// TIA Portal V21 export
FUNCTION_BLOCK "FB_StarterStl"   // FB103, STL
TITLE = Пускатель насоса (STL)
{ S7_Optimized_Access := 'FALSE' }
AUTHOR : WTP2
FAMILY : Drives
VERSION : 0.1
// Пускатель насоса с контролем обратной связи (один блок на LAD, FBD, STL, SCL).
// 1. Пуск/стоп — SR с битом-операндом xRunMem: S = xStart AND xInterlock; R1 = xStop OR NOT xInterlock OR xFault.
//    SR S7: сначала S, затем R1 — при S = R1 = 1 (Пуск и Стоп одновременно) бит сброшен. xRun := xRunMem.
// 2. Контроль обратной связи: TON tonFeedback (IN = xRun AND NOT xFeedback, PT = tFeedbackTime).
// 3. Авария с самоподхватом: xFault := (tonFeedback.Q OR xFault) AND NOT xReset.
// 4. Счётчик пусков: по фронту xRun (бит памяти xEdgeMem) iStarts := iStarts + 1.
// Порядок сетей 1-4; xFault в сети 1 — значение прошлого вызова.
// stored: AutoNumber false, SetENOAutomatically false
   VAR_INPUT
      xStart : Bool;   // Пуск (кнопка)
      xStop : Bool;   // Стоп (кнопка, TRUE — нажата)
      xInterlock : Bool := TRUE;   // Блокировки в норме, пуск разрешён
      xFeedback : Bool;   // Обратная связь контактора
      tFeedbackTime : Time := T#2S;   // Допустимое время без обратной связи
      xReset : Bool;   // Сброс аварии
   END_VAR
   VAR_OUTPUT
      xRun : Bool;   // Команда контактору
      xFault : Bool;   // Авария: нет обратной связи
      iStarts : Int;   // Число пусков
   END_VAR
   VAR
      xRunMem : Bool;   // Бит-операнд SR пуска
      xEdgeMem : Bool;   // Бит памяти фронта xRun
      tonFeedback : TON_TIME;   // Таймер контроля обратной связи
   END_VAR
   VAR_TEMP
      xTonIn : Bool;   // Вход таймера
      xTonQ : Bool;   // Выход таймера
   END_VAR
BEGIN

NETWORK
TITLE = Пуск/стоп: SR, сброс главнее
      A     #xStart;
      A     #xInterlock;
      S     #xRunMem;
      A     #xStop;
      ON    #xInterlock;
      O     #xFault;
      R     #xRunMem;
      A     #xRunMem;
      =     #xRun;

NETWORK
TITLE = Контроль обратной связи
      A     #xRun;
      AN    #xFeedback;
      =     #xTonIn;
      CALL  #tonFeedback
      ( IN := #xTonIn,
        PT := #tFeedbackTime,
        Q  := #xTonQ,
        ET := 
      );

NETWORK
TITLE = Авария с самоподхватом
      A(;
      O     #xTonQ;
      O     #xFault;
      );
      AN    #xReset;
      =     #xFault;

NETWORK
TITLE = Счётчик пусков по фронту xRun
      A     #xRun;
      FP    #xEdgeMem;
      JCN   M001;
      L     #iStarts;
      L     1;
      +I;
      T     #iStarts;
M001: NOP   0;
END_FUNCTION_BLOCK
